SUBAPPLICATION Uebung_259b_AX (* Gamma mit Rampe, Taster: I1 = 0, I2 = 4000, I3 = 8000, I4 = 2000 auf LED Q1 linear und LED Q2 Gamma 2.2, beide RAMP 2s *)
  (* Standard: 61499-2; Description: Copyright (c) 2026 Meisterschulen am Ostbahnhof This program and the accompanying materials are made available under the terms of the Eclipse Public License 2.0 which is available at https://www.eclipse.org/legal/epl-2.0/ SPDX-License-Identifier: EPL-2.0 *)
  (* Version 1.0, 2026-11-06, Franz Höpfinger, Meisterschulen am Ostbahnhof, initial API and implementation and/or initial documentation *)
  PACKAGE Uebungen;
  IMPORT logiBUS::io::DI::logiBUS_DI::Input_I1;
  IMPORT logiBUS::io::DI::logiBUS_DI::Input_I2;
  IMPORT logiBUS::io::DI::logiBUS_DI::Input_I3;
  IMPORT logiBUS::io::DI::logiBUS_DI::Input_I4;
  IMPORT logiBUS::io::DI::logiBUS_DI_Events::BUTTON_PRESS_DOWN;
  IMPORT logiBUS::io::DQ::logiBUS_DO::Output_Q1;
  IMPORT logiBUS::io::DQ::logiBUS_DO::Output_Q2;
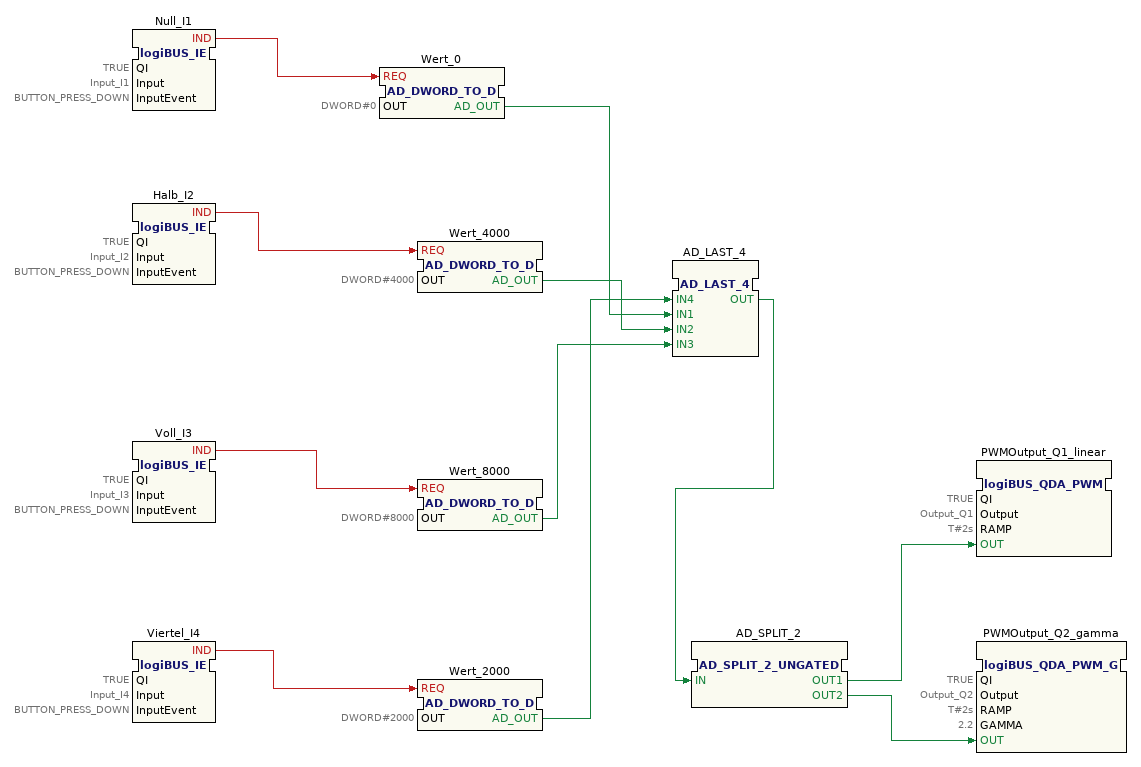
  FBS
    Null_I1 : logiBUS::io::DI::logiBUS_IE(QI := TRUE, Input := Input_I1, InputEvent := BUTTON_PRESS_DOWN);
    Wert_0 : adapter::conversion::unidirectional::AD_DWORD_TO_D(OUT := DWORD#0);
    Halb_I2 : logiBUS::io::DI::logiBUS_IE(QI := TRUE, Input := Input_I2, InputEvent := BUTTON_PRESS_DOWN);
    Wert_4000 : adapter::conversion::unidirectional::AD_DWORD_TO_D(OUT := DWORD#4000);
    Voll_I3 : logiBUS::io::DI::logiBUS_IE(QI := TRUE, Input := Input_I3, InputEvent := BUTTON_PRESS_DOWN);
    Wert_8000 : adapter::conversion::unidirectional::AD_DWORD_TO_D(OUT := DWORD#8000);
    Viertel_I4 : logiBUS::io::DI::logiBUS_IE(QI := TRUE, Input := Input_I4, InputEvent := BUTTON_PRESS_DOWN);
    Wert_2000 : adapter::conversion::unidirectional::AD_DWORD_TO_D(OUT := DWORD#2000);
    AD_LAST_4 : adapter::events::unidirectional::AD_LAST_4;
    AD_SPLIT_2 : adapter::events::unidirectional::AD_SPLIT_2_UNGATED;
    PWMOutput_Q1_linear : logiBUS::io::DQ::logiBUS_QDA_PWM(QI := TRUE, Output := Output_Q1, RAMP := T#2s);
    PWMOutput_Q2_gamma : logiBUS::io::DQ::logiBUS_QDA_PWM_G(QI := TRUE, Output := Output_Q2, RAMP := T#2s, GAMMA := 2.2);
  END_FBS
  EVENT_CONNECTIONS
    Viertel_I4.IND TO Wert_2000.REQ;
    Null_I1.IND TO Wert_0.REQ;
    Halb_I2.IND TO Wert_4000.REQ;
    Voll_I3.IND TO Wert_8000.REQ;
  END_CONNECTIONS
  ADAPTER_CONNECTIONS
    Wert_2000.AD_OUT TO AD_LAST_4.IN4;
    Wert_0.AD_OUT TO AD_LAST_4.IN1;
    Wert_4000.AD_OUT TO AD_LAST_4.IN2;
    Wert_8000.AD_OUT TO AD_LAST_4.IN3;
    AD_LAST_4.OUT TO AD_SPLIT_2.IN;
    AD_SPLIT_2.OUT1 TO PWMOutput_Q1_linear.OUT;
    AD_SPLIT_2.OUT2 TO PWMOutput_Q2_gamma.OUT;
  END_CONNECTIONS
END_SUBAPPLICATION
